// TIA Portal project "LAB06" (V16)

(* hardware
DEVICE "S7300/ET200M station_1"  S7-300 station
   slot 0: "Rail_0"  Rail  6ES7 390-1***0-0AA0
   slot 2: "PLC_1"  CPU 313C-2 DP  6ES7 313-6CF03-0AB0  V2.6
      slot 0: "MPI interface_1"  X1
      slot 1: "DP interface_1"  X2
      slot 2: "DI 16/DO 16_1"  DI16/DO16
      slot 4: "Count_1"  Counter
*)

// ===== PLC "PLC_1"  CPU 313C-2 DP =====

VAR_GLOBAL   // PLC tag table "Default tag table"
   "Tag_1" AT %MW0 : Word;
   "Tag_2" AT %MW2 : Word;
   "Tag_3" AT %MW4 : Word;
   "Tag_4" AT %MW6 : Word;
   "Tag_5" AT %MD8 : DWord;
   "Tag_6" AT %MW12 : Word;
   "Tag_7" AT %MW20 : Word;
   "Tag_8" AT %MW22 : Int;
   "Tag_9" AT %M20.0 : Bool;
   "Tag_10" AT %MB20 : Byte;
   "Tag_11" AT %MW24 : Int;
   "Tag_12" AT %MD14 : DWord;
   "Tag_13" AT %MW8 : Word;
   "Tag_14" AT %M26.0 : Bool;
   "Tag_15" AT %MW28 : Int;
   "Tag_16" AT %MW16 : Word;
   "Tag_17" AT %MW18 : Word;
END_VAR

DATA_BLOCK "DB100"   // DB100
{ S7_Optimized_Access := 'FALSE' }
VERSION : 0.1
   VAR
      Static_1 : Int := 10;
      Static_2 : Int := 20;
      Static_3 : Int := 30;
      Static_4 : Int := 40;
   END_VAR
BEGIN
END_DATA_BLOCK

DATA_BLOCK "DB101"   // DB101
{ S7_Optimized_Access := 'FALSE' }
VERSION : 0.1
   VAR
      Static_1 : Int := 99;
      Static_2 : Int := 99;
      Static_3 : Int := 99;
      Static_4 : Int := 99;
      Static_5 : Int := 99;
      Static_6 : Int := 0;
      Static_7 : Int;
      Static_8 : Int;
      Static_9 : Int;
   END_VAR
BEGIN
END_DATA_BLOCK

FUNCTION "FC8" : Void   // FC8, STL
{ S7_Optimized_Access := 'FALSE' }
VERSION : 0.1
   VAR_INPUT
      db_source : Int;
      db_destination : Int;
   END_VAR
   VAR_OUTPUT
      error : Bool;
      length : Int;
   END_VAR
BEGIN

REGION Network 1
   // vars inizialization
         L     0;  // reset output parameter length
         T     #length;
         CLR;  // instruction that puts RLO=0
         =     #error;  // error parameter initialized to 0
   // DB source
         L     #db_source;  // load number of db source
         T     "Tag_1";
         OPN   DB["Tag_1"];  // indirect opening of db source
         L     DBLG;
         T     "Tag_2";  // save length in MW2
   // DB destination
         L     #db_destination;  // load number of db destination
         T     "Tag_3";
         OPN   DB["Tag_3"];  // indirect opening of db destination
         L     DBLG;
         T     "Tag_4";  // save length in MW6
   // length check
         L     "Tag_2";  // load length of db source
         <I;  // if destination length < source length
         =     #error;  // error parameter =1
         BEC;  // return
   // transfer allowed
         L     P#0.0;  // else proceed with db transfer
         T     "Tag_5";  // initialize pointer for data blocks
         L     "Tag_2";  // load length of db source
         T     #length;  // calculation of the number of iterations
         L     2;
         /I;

   TRAF: T     "Tag_6";  // save on MW12
         OPN   DB["Tag_1"];  // open db source
         L     DBW [ "Tag_5"];  // load word of db source
         OPN   DB["Tag_3"];  // open db destination
         T     DBW [ "Tag_5"];  // transfer in db destination
         L     P#2.0;
         L     "Tag_5";  // increment pointer
         +D;
         T     "Tag_5";
         L     "Tag_6";  // load number of iterations
         LOOP  TRAF;
END_REGION
END_FUNCTION

FUNCTION "FC81" : Void   // FC81, STL
{ S7_Optimized_Access := 'FALSE' }
VERSION : 0.1
   VAR_INPUT
      db_source : Int;
      db_destination : Int;
   END_VAR
   VAR_OUTPUT
      error : Int;
      length : Int;
   END_VAR
BEGIN

REGION Network 1
   // vars inizialization
         L     0;  // reset output parameter length
         T     #length;
         L     0;
         T     #error;  // error parameter initialized to 0
   // DB source
         L     #db_source;  // load number of db source
         T     "Tag_1";
         OPN   DB["Tag_1"];  // indirect opening of db source
         L     DBLG;
         T     "Tag_2";  // save length in MW2
   // DB destination
         L     #db_destination;  // load number of db destination
         T     "Tag_3";
         OPN   DB["Tag_3"];  // indirect opening of db destination
         L     DBLG;
         T     "Tag_4";  // save length in MW6
   // length check
         L     "Tag_2";  // load length of db source
         <I;  // if destination length < source length
         JCN   OK;  // if we have enough space, jump to OK
         L     -1;
         T     #error;  // error parameter = -1
         L     "Tag_4";  // overwrite MW2 with destination length
         T     "Tag_2";
   OK:   NOP   0;

   // transfer allowed
         L     P#0.0;  // else proceed with db transfer
         T     "Tag_5";  // initialize pointer for data blocks
         L     "Tag_2";  // load length of db source
         T     #length;  // calculation of the number of iterations
         L     2;
         /I;

   TRAF: T     "Tag_6";  // save on MW12
         OPN   DB["Tag_1"];  // open db source
         L     DBW [ "Tag_5"];  // load word of db source
         OPN   DB [ "Tag_3"];  // open db destination
         T     DBW [ "Tag_5"];  // transfer in db destination
         L     P#2.0;
         L     "Tag_5";  // increment pointer
         +D;
         T     "Tag_5";
         L     "Tag_6";  // load number of iterations
         LOOP  TRAF;
END_REGION
END_FUNCTION

FUNCTION "FC82" : Void   // FC82, STL
{ S7_Optimized_Access := 'FALSE' }
VERSION : 0.1
   VAR_INPUT
      db_source : Int;
      db_destination : Int;
   END_VAR
   VAR_OUTPUT
      error : Bool;
      length : Int;
   END_VAR
BEGIN

REGION Network 1
   // vars inizialization
         L     0;  // reset output parameter length
         T     #length;
         CLR;  // instruction that puts RLO=0
         =     #error;  // error parameter initialized to 0
   // DB source
         L     #db_source;  // load number of db source
         T     "Tag_1";
         OPN   DB["Tag_1"];  // indirect opening of db source
         L     DBLG;
         T     "Tag_2";  // save length in MW2
   // DB destination
         L     #db_destination;  // load number of db destination
         T     "Tag_3";
         OPN   DB["Tag_3"];  // indirect opening of db destination
         L     DBLG;
         T     "Tag_4";  // save length in MW6
   // length check
         L     "Tag_2";  // load length of db source
         L     10;
         +I;  // source + 10
         T     "Tag_17";  // saves (source + 10) in MW18

         L     "Tag_4";  // load length of db destination
         L     "Tag_17";
         <I;  // if destination length < (source + 10)
         =     #error;  // error parameter =1
         BEC;  // return
   // transfer allowed
         L     P#0.0;  // else proceed with db transfer
         T     "Tag_5";  // initialize pointer for data blocks
         L     "Tag_2";  // load length of db source
         T     #length;  // calculation of the number of iterations
         L     2;
         /I;

   TRAF: T     "Tag_6";  // save on MW12
         L     "Tag_5";  // compute MD14 = MD8 + 10 bytes
         L     P#10.0;
         +D;
         T     "Tag_12";

         OPN   DB["Tag_1"];  // open db source
         L     DBW [ "Tag_5"];  // load word of db source
         OPN   DB["Tag_3"];  // open db destination
         T     DBW [ "Tag_12"];  // transfer in db destination

         L     P#2.0;
         L     "Tag_5";  // increment pointer
         +D;
         T     "Tag_5";  // update MD8
         L     "Tag_6";  // load number of iterations
         LOOP  TRAF;
END_REGION
END_FUNCTION

ORGANIZATION_BLOCK "Main"   // OB1, STL
TITLE = "Main Program Sweep (Cycle)"
{ S7_Optimized_Access := 'FALSE' }
VERSION : 0.1
   VAR_TEMP
      OB1_EV_CLASS : Byte;   // Bits 0-3 = 1 (Coming event), Bits 4-7 = 1 (Event class 1)
      OB1_SCAN_1 : Byte;   // 1 (Cold restart scan 1 of OB 1), 3 (Scan 2-n of OB 1)
      OB1_PRIORITY : Byte;   // Priority of OB Execution
      OB1_OB_NUMBR : Byte;   // 1 (Organization block 1, OB1)
      OB1_RESERVED_1 : Byte;   // Reserved for system
      OB1_RESERVED_2 : Byte;   // Reserved for system
      OB1_PREV_CYCLE : Int;   // Cycle time of previous OB1 scan (milliseconds)
      OB1_MIN_CYCLE : Int;   // Minimum cycle time of OB1 (milliseconds)
      OB1_MAX_CYCLE : Int;   // Maximum cycle time of OB1 (milliseconds)
      OB1_DATE_TIME : Date_And_Time;   // Date and time OB1 started
   END_VAR
BEGIN

REGION Network 1
         CALL  "FC82"
         ( db_source      := 100,
           db_destination := 101,
           error          := "Tag_14",
           length         := "Tag_15"
         );
END_REGION
END_ORGANIZATION_BLOCK